(* IEC 61131-3 sources: rusty/tests/lit/cfc/generics/generic_feedback, 2 files *)

(* ---- main.st ---- *)
FUNCTION main : DINT
    generic_feedback.seed := 5;
    generic_feedback();
    generic_feedback();
    generic_feedback();
    // CHECK: acc = 15
    printf('acc = %d$N', generic_feedback.acc);
END_FUNCTION

(* ---- myGenAdd.st ---- *)
FUNCTION myGenAdd<T: ANY_NUM> : T
VAR_INPUT
    a : T;
    b : T;
END_VAR
END_FUNCTION

FUNCTION myGenAdd__DINT : DINT
VAR_INPUT
    a : DINT;
    b : DINT;
END_VAR
    myGenAdd__DINT := a + b;
END_FUNCTION
